Staubli VAL3: toolItem.dtx

public string sName
public tool tTool = {fatherId=flange[0]}
